FUNCTION_BLOCK TransportGeneral1 (* CAT Function Block Type *)
  (* Standard: 61499-2 *)
  (* Version 0.0, 7/10/2026, template *)
  PACKAGE Main;
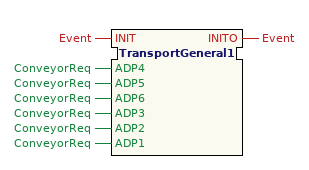
  EVENT_INPUT
    INIT; (* Initialization Request *)
  END_EVENT
  EVENT_OUTPUT
    INITO; (* Initialization Confirm *)
  END_EVENT
  SOCKETS
    ADP4 : ConveyorReq;
    ADP5 : ConveyorReq;
    ADP6 : ConveyorReq;
    ADP3 : ConveyorReq;
    ADP2 : ConveyorReq;
    ADP1 : ConveyorReq;
  END_SOCKETS
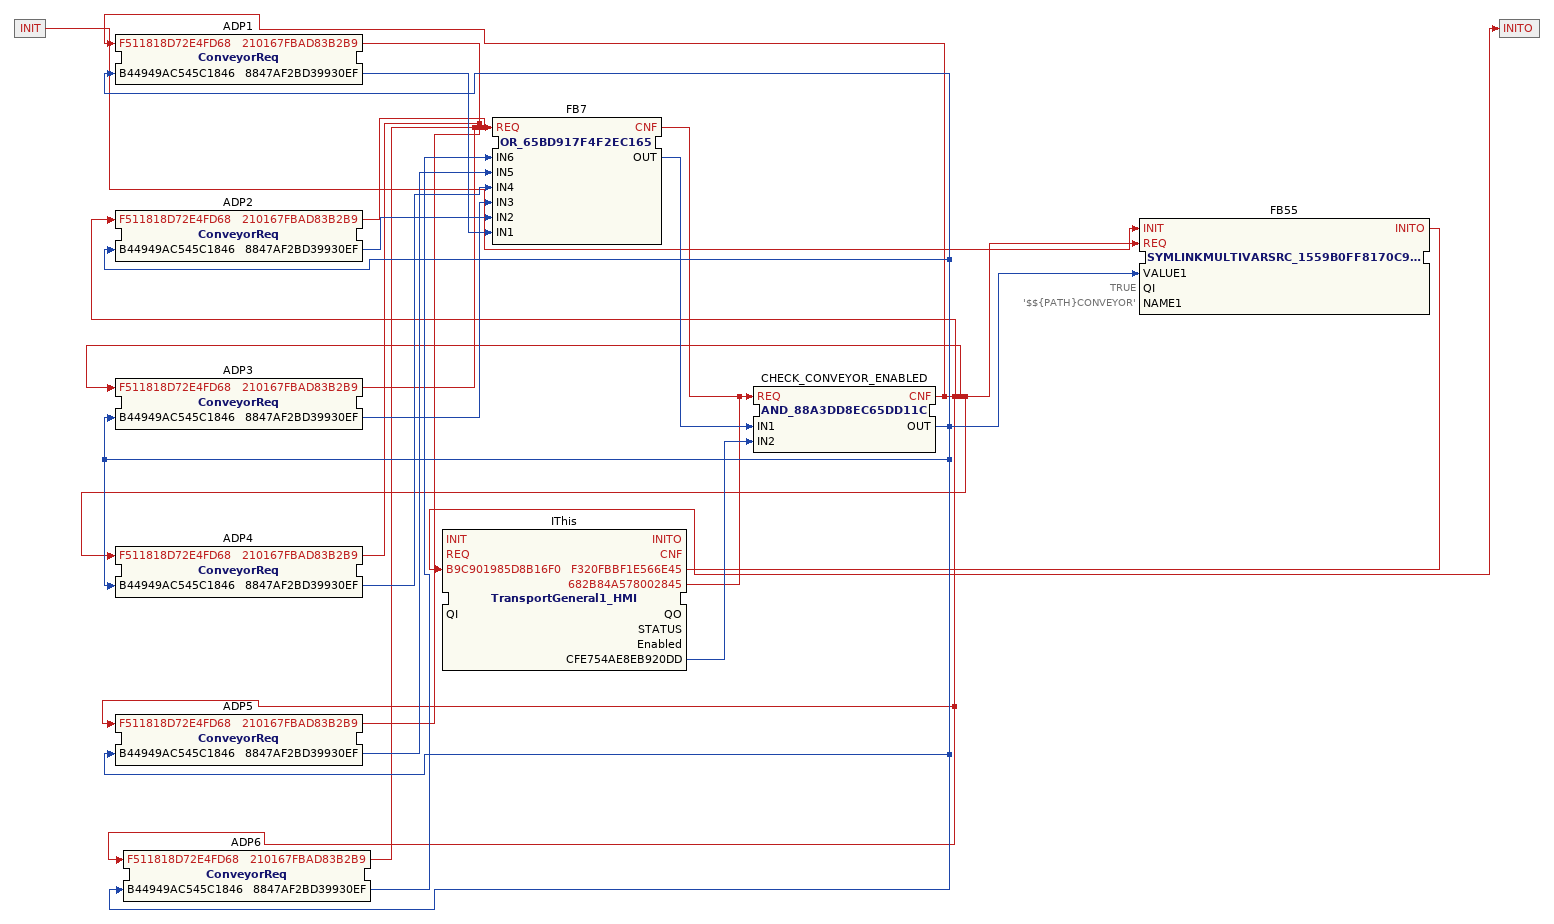
  FBS
    FB7 : OR_65BD917F4F2EC165; {SET_ATTRIBUTE(Configuration.GenericFBType.InterfaceParams, Runtime.Standard#CNT:=6;OUT:BOOL)}
    IThis : TransportGeneral1_HMI;
    CHECK_CONVEYOR_ENABLED : AND_88A3DD8EC65DD11C; {SET_ATTRIBUTE(Configuration.GenericFBType.InterfaceParams, Runtime.Standard#CNT:=2;OUT:BOOL)}
    FB55 : SYMLINKMULTIVARSRC_1559B0FF8170C9BA0(QI := TRUE, NAME1 := '$${PATH}CONVEYOR'); {SET_ATTRIBUTE(Configuration.GenericFBType.InterfaceParams, Runtime.System#I:=1;VALUE${I$}:BOOL)}
  END_FBS
  EVENT_CONNECTIONS
    FB7.CNF TO CHECK_CONVEYOR_ENABLED.REQ;
    INIT TO FB55.INIT;
    CHECK_CONVEYOR_ENABLED.CNF TO FB55.REQ;
    ADP6.210167FBAD83B2B9 TO FB7.REQ;
    ADP5.210167FBAD83B2B9 TO FB7.REQ;
    ADP4.210167FBAD83B2B9 TO FB7.REQ;
    FB55.INITO TO IThis.B9C901985D8B16F0;
    IThis.F320FBBF1E566E45 TO INITO;
    IThis.682B84A578002845 TO CHECK_CONVEYOR_ENABLED.REQ;
    ADP3.210167FBAD83B2B9 TO FB7.REQ;
    ADP2.210167FBAD83B2B9 TO FB7.REQ;
    ADP1.210167FBAD83B2B9 TO FB7.REQ;
    CHECK_CONVEYOR_ENABLED.CNF TO ADP1.F511818D72E4FD68;
    CHECK_CONVEYOR_ENABLED.CNF TO ADP2.F511818D72E4FD68;
    CHECK_CONVEYOR_ENABLED.CNF TO ADP3.F511818D72E4FD68;
    CHECK_CONVEYOR_ENABLED.CNF TO ADP4.F511818D72E4FD68;
    CHECK_CONVEYOR_ENABLED.CNF TO ADP5.F511818D72E4FD68;
    CHECK_CONVEYOR_ENABLED.CNF TO ADP6.F511818D72E4FD68;
  END_CONNECTIONS
  DATA_CONNECTIONS
    CHECK_CONVEYOR_ENABLED.OUT TO FB55.VALUE1;
    FB7.OUT TO CHECK_CONVEYOR_ENABLED.IN1;
    ADP6.8847AF2BD39930EF TO FB7.IN6;
    ADP5.8847AF2BD39930EF TO FB7.IN5;
    ADP4.8847AF2BD39930EF TO FB7.IN4;
    IThis.CFE754AE8EB920DD TO CHECK_CONVEYOR_ENABLED.IN2;
    ADP3.8847AF2BD39930EF TO FB7.IN3;
    ADP2.8847AF2BD39930EF TO FB7.IN2;
    ADP1.8847AF2BD39930EF TO FB7.IN1;
    CHECK_CONVEYOR_ENABLED.OUT TO ADP1.B44949AC545C1846;
    CHECK_CONVEYOR_ENABLED.OUT TO ADP2.B44949AC545C1846;
    CHECK_CONVEYOR_ENABLED.OUT TO ADP3.B44949AC545C1846;
    CHECK_CONVEYOR_ENABLED.OUT TO ADP4.B44949AC545C1846;
    CHECK_CONVEYOR_ENABLED.OUT TO ADP5.B44949AC545C1846;
    CHECK_CONVEYOR_ENABLED.OUT TO ADP6.B44949AC545C1846;
  END_CONNECTIONS
END_FUNCTION_BLOCK
